# B&R Automation Studio project DemoCNC (part 2)

#### Variables.var - Local variables
```iecst
VAR
	deviceName : STRING[20] := 'CNC_PrgDir'; (*file device of the CNC programs (FileDevice of the axes group program feature, Config_4)*)
	shareParam : STRING[200] := '/SIP=192.0.2.20 /PROTOCOL=cifs /SHARE=GCode /USER=Controller /PASSWORD=change-me'; (*network share holding the CNC programs (HMI PC) - example values : set the address and the account of your PC*)
	step : USINT := 0;
	fbDevLink : DevLink;
	retryTimer : TON;
	linked : BOOL := FALSE; (*TRUE = the program folder is available*)
	linkStatus : UINT := 0; (*status of the last failed link, 0 = none*)
	sysError : UDINT := 0; (*FileIoGetSysError of the last failed link*)
END_VAR
```

### Package Logical/Motion - Manual axis moves, handwheel, path trace

### Program Logical/Motion/AxisManual (IEC) - Manual axis moves : jog, position move, single-axis commands

#### Init.st - Init code
```iecst
PROGRAM _INIT

	gEquipment.Output.Status.MoveComplete := TRUE;

	FOR i := 0 TO AX_LAST DO
		gAxis[i].Input.Parameter.JogSpeed := 50;
	END_FOR;

	(* static axis references : index 0 = X, 1 = Y, 2 = Z *)
	fbAxisInfo[AX_X].Axis := ADR(gAxis_X);
	fbAxisInfo[AX_Y].Axis := ADR(gAxis_Y);
	fbAxisInfo[AX_Z].Axis := ADR(gAxis_Z);

	fbAxisStatus[AX_X].Axis := ADR(gAxis_X);
	fbAxisStatus[AX_Y].Axis := ADR(gAxis_Y);
	fbAxisStatus[AX_Z].Axis := ADR(gAxis_Z);

	fbAxisPosition[AX_X].Axis := ADR(gAxis_X);
	fbAxisPosition[AX_Y].Axis := ADR(gAxis_Y);
	fbAxisPosition[AX_Z].Axis := ADR(gAxis_Z);

	fbAxisVelocity[AX_X].Axis := ADR(gAxis_X);
	fbAxisVelocity[AX_Y].Axis := ADR(gAxis_Y);
	fbAxisVelocity[AX_Z].Axis := ADR(gAxis_Z);

	fbAxisTorque[AX_X].Axis := ADR(gAxis_X);
	fbAxisTorque[AX_Y].Axis := ADR(gAxis_Y);
	fbAxisTorque[AX_Z].Axis := ADR(gAxis_Z);

	fbMoveAbs[AX_X].Axis := ADR(gAxis_X);
	fbMoveAbs[AX_Y].Axis := ADR(gAxis_Y);
	fbMoveAbs[AX_Z].Axis := ADR(gAxis_Z);

	fbMoveAdd[AX_X].Axis := ADR(gAxis_X);
	fbMoveAdd[AX_Y].Axis := ADR(gAxis_Y);
	fbMoveAdd[AX_Z].Axis := ADR(gAxis_Z);

	fbJog[AX_X].Axis := ADR(gAxis_X);
	fbJog[AX_Y].Axis := ADR(gAxis_Y);
	fbJog[AX_Z].Axis := ADR(gAxis_Z);

	fbStop[AX_X].Axis := ADR(gAxis_X);
	fbStop[AX_Y].Axis := ADR(gAxis_Y);
	fbStop[AX_Z].Axis := ADR(gAxis_Z);

	fbHalt[AX_X].Axis := ADR(gAxis_X);
	fbHalt[AX_Y].Axis := ADR(gAxis_Y);
	fbHalt[AX_Z].Axis := ADR(gAxis_Z);

	fbReset[AX_X].Axis := ADR(gAxis_X);
	fbReset[AX_Y].Axis := ADR(gAxis_Y);
	fbReset[AX_Z].Axis := ADR(gAxis_Z);

	fbAxisError[AX_X].Axis := ADR(gAxis_X);
	fbAxisError[AX_Y].Axis := ADR(gAxis_Y);
	fbAxisError[AX_Z].Axis := ADR(gAxis_Z);

	fbPower[AX_X].Axis := ADR(gAxis_X);
	fbPower[AX_Y].Axis := ADR(gAxis_Y);
	fbPower[AX_Z].Axis := ADR(gAxis_Z);

	fbHome[AX_X].Axis := ADR(gAxis_X);
	fbHome[AX_Y].Axis := ADR(gAxis_Y);
	fbHome[AX_Z].Axis := ADR(gAxis_Z);

	FOR i := 0 TO AX_LAST DO
		fbAxisInfo[i].Enable := TRUE;
		fbAxisStatus[i].Enable := TRUE;
		fbAxisPosition[i].Enable := TRUE;
		fbAxisVelocity[i].Enable := TRUE;
		fbAxisTorque[i].Enable := TRUE;
		fbAxisError[i].Enable := TRUE;

		fbJog[i].Acceleration := DEFAULT_ACC;
		fbJog[i].Deceleration := DEFAULT_DEC;
		fbMoveAbs[i].Acceleration := DEFAULT_ACC;
		fbMoveAbs[i].Deceleration := DEFAULT_DEC;
		fbMoveAdd[i].Acceleration := DEFAULT_ACC;
		fbMoveAdd[i].Deceleration := DEFAULT_DEC;
		fbStop[i].Deceleration := DEFAULT_DEC;
		fbHalt[i].Deceleration := DEFAULT_DEC;
	END_FOR

END_PROGRAM
```

#### Cyclic.st - Cyclic code
```iecst
PROGRAM _CYCLIC

	(* drive adapter PVs (Global.var) : referenced here so they are allocated on the target *)
	gDS402_X;
	gDS402_Y;
	gDS402_Z;

	(* copy the mappMotion position limits into gAxis[].Input.Parameter.SoftwareLimits* once after startup *)
	IF NOT cfgLimitLoaded THEN
		fbAxCfg.Name := cfgAxisName[cfgAxIdx];
		fbAxCfg.DataType := mcCFG_AX_MOVE_LIM;
		fbAxCfg.DataAddress := ADR(axMoveLim);
		fbAxCfg.Mode := mcPCM_LOAD;
		fbAxCfg.Execute := TRUE;
		fbAxCfg();

		IF fbAxCfg.Done OR fbAxCfg.Error THEN
			cfgLimitErrorID[cfgAxIdx] := fbAxCfg.ErrorID;
			IF fbAxCfg.Done THEN
				gAxis[cfgAxIdx].Input.Parameter.SoftwareLimitsNeg := LREAL_TO_DINT(axMoveLim.MovementLimits.Internal.Position.LowerLimit);
				gAxis[cfgAxIdx].Input.Parameter.SoftwareLimitsPos := LREAL_TO_DINT(axMoveLim.MovementLimits.Internal.Position.UpperLimit);
			END_IF
			fbAxCfg.Execute := FALSE;
			fbAxCfg();
			cfgAxIdx := cfgAxIdx + 1;
			cfgLimitLoaded := cfgAxIdx > AX_LAST;
		END_IF
	END_IF

	Torque_X := fbAxisTorque[AX_X].Torque;
	Torque_Y := fbAxisTorque[AX_Y].Torque;
	Torque_Z := fbAxisTorque[AX_Z].Torque;

	(* absolute positions are meaningless before homing *)
	allHomed := fbAxisInfo[AX_X].IsHomed AND fbAxisInfo[AX_Y].IsHomed AND fbAxisInfo[AX_Z].IsHomed;

	(* position move request of this scan : accepted or dropped below, reported by act_MoveResult *)
	moveReq := gEquipment.Input.Command.ManualMove;
	moveAccepted := FALSE;

	IF NOT DI_MPG_Jog_Enable AND gEquipment.Input.CncCommand = E_ACT_IDLE AND NOT gEquipment.Output.State.Move AND NOT DI_Auto AND NOT gEquipment.Output.Status.EmergencyStop THEN

		IF NOT allHomed THEN
			gEquipment.Input.Command.ManualMove := FALSE;
		END_IF

		IF gEquipment.Input.Command.ManualMove THEN
			gEquipment.Input.Command.ManualMove := FALSE;
			gEquipment.Output.Status.MoveComplete := FALSE;
			moveStep := 0;
			moveAccepted := TRUE;
		END_IF

		act_Jog;
	ELSE
		gEquipment.Output.Status.ManualMove := FALSE;
		gEquipment.Input.Command.ManualMove := FALSE; (* never run a stale move request later *)
	END_IF

	moveStepIn := moveStep;
	act_MovePosition;
	act_MoveResult; (* result to the HMI (gManualMoveResult) - reporting only *)

	(* per-axis POWER / HOME only while the CNC is idle *)
	cncIdle := gEquipment.Output.Status.CurrentAction = E_ACT_IDLE AND NOT gEquipment.Output.Status.ProgramActive;

	(* screen jog (Axis_JOG_POSITIVE / NEGATIVE) only in manual mode, without the handwheel and while no CNC command runs.
	   MOVE_ADDITIVE (one step) is not gated : the HMI uses it in auto mode too.
	   Not ProgramActive (cncIdle) : the axes group reports MoveActive for a cycle when a single axis starts to move, so every
	   jog would be dropped right after its start. A program only runs in auto mode, which NOT DI_Auto already keeps out *)
	jogAllowed := NOT DI_Auto AND NOT DI_MPG_Jog_Enable AND gEquipment.Output.Status.CurrentAction = E_ACT_IDLE;

	(* per-axis power is held by fbPower (Axis_POWER). E-stop and group servo off take the axes back *)
	IF gEquipment.Output.Status.EmergencyStop OR gEquipment.Output.Status.CurrentAction = E_ACT_POWER_OFF THEN
		FOR i := 0 TO AX_LAST BY 1 DO
			axisPowerReq[i] := FALSE;
		END_FOR
	END_IF

	(* jog watchdog : an HMI that changes gJogAlive while it jogs (every 0.1 s) gets the jog stopped when the value
	   stands still for 0.5 s (HMI hung, connection lost). An HMI that never changes it is not watched *)
	jogAny := jogPosActive[AX_X] OR jogNegActive[AX_X] OR jogPosActive[AX_Y] OR jogNegActive[AX_Y] OR jogPosActive[AX_Z] OR jogNegActive[AX_Z];
	IF NOT jogAny THEN
		jogAliveArmed := FALSE;
		jogAlivePrev := gJogAlive;
	ELSIF gJogAlive <> jogAlivePrev THEN
		jogAlivePrev := gJogAlive;
		jogAliveArmed := TRUE;
		jogAliveTimer(IN := FALSE); (* restart *)
	END_IF
	jogAliveTimer(IN := jogAny AND jogAliveArmed, PT := T#500ms);
	IF jogAliveTimer.Q THEN
		FOR i := 0 TO AX_LAST BY 1 DO
			jogPosActive[i] := FALSE;
			jogNegActive[i] := FALSE;
		END_FOR
		jogAliveArmed := FALSE;
	END_IF

	(* ---------- per-axis command handling ---------- *)
	FOR i := 0 TO AX_LAST BY 1 DO

		(* E-stop : stop whatever runs, accept only STOP / RESET *)
		IF gEquipment.Output.Status.EmergencyStop THEN
			IF gAxis[i].Input.Command.Command <> Axis_STOP AND gAxis[i].Input.Command.Command <> Axis_RESET THEN
				gAxis[i].Input.Command.Command := Axis_IDLE;
			END_IF
			IF (command[i] <> Axis_IDLE AND command[i] <> Axis_STOP AND command[i] <> Axis_RESET) OR jogPosActive[i] OR jogNegActive[i] THEN
				command[i] := Axis_STOP;
				commandStep[i] := 0;
			END_IF
		END_IF

		IF command[i] <> gAxis[i].Input.Command.Command AND command[i] = Axis_IDLE THEN
			gAxis[i].Output.State.Command := gAxis[i].Input.Command.Command;
			command[i] := gAxis[i].Input.Command.Command;
			gAxis[i].Input.Command.Command := Axis_IDLE;
			commandStep[i] := 0;
		ELSIF gAxis[i].Input.Command.Command = Axis_HALT AND command[i] <> Axis_IDLE THEN
			command[i] := gAxis[i].Input.Command.Command;
			gAxis[i].Input.Command.Command := Axis_IDLE;
			commandStep[i] := 0;
		ELSIF gAxis[i].Input.Command.Command = Axis_STOP AND command[i] <> Axis_IDLE THEN
			command[i] := gAxis[i].Input.Command.Command;
			gAxis[i].Input.Command.Command := Axis_IDLE;
			commandStep[i] := 0;
		END_IF

		(* a HALT / STOP ends a running position move (act_MovePosition never sends them itself) *)
		IF (command[i] = Axis_HALT OR command[i] = Axis_STOP) AND commandStep[i] = 0 AND moveStep < 100 THEN
			moveStep := 100;
		END_IF

		CASE command[i] OF
			Axis_IDLE:
				IF fbAxisInfo[i].IsHomed THEN
					gAxis[i].Output.State.Status := 1;
				ELSE
					gAxis[i].Output.State.Status := 0;
				END_IF

				gAxis[i].Output.State.Home := fbAxisInfo[i].IsHomed;

				(* keep jog active state while jogging (command returns to IDLE, motion continues) *)
				IF jogPosActive[i] OR jogNegActive[i] THEN
					gAxis[i].Output.State.Status := 2;
				END_IF

			Axis_HALT:
				CASE commandStep[i] OF
					0:
						IF (jogPosActive[i] OR jogNegActive[i]) AND NOT fbMoveAbs[i].Busy AND NOT fbMoveAdd[i].Busy AND NOT fbHome[i].Busy THEN
							(* jog only : the jog FB brakes by itself (Deceleration) when its request drops. MC_Halt would abort it,
							   and an aborted jog FB took no new jog until it was switched off and on *)
							jogPosActive[i] := FALSE;
							jogNegActive[i] := FALSE;
							fbMoveAbs[i].Execute := FALSE; (* not busy - released as in the MC_Halt path *)
							fbMoveAdd[i].Execute := FALSE;
							fbHome[i].Execute := FALSE;
							settleTimer[i](IN := FALSE);
							commandStep[i] := 2;
						ELSE
							jogPosActive[i] := FALSE;
							jogNegActive[i] := FALSE;
							fbMoveAbs[i].Execute := FALSE; (* release aborted moves so the next one gets a rising edge *)
							fbMoveAdd[i].Execute := FALSE;
							fbHome[i].Execute := FALSE;
							fbHalt[i].Execute := TRUE;
							settleTimer[i](IN := FALSE);
							commandStep[i] := 1;
						END_IF
					1:
						IF fbHalt[i].Done OR fbHalt[i].CommandAborted OR fbHalt[i].Error THEN
							fbHalt[i].Execute := FALSE;
							IF fbAxisStatus[i].StandStill OR fbAxisStatus[i].ErrorStop OR fbAxisStatus[i].Disabled THEN
								command[i] := Axis_IDLE;
							ELSE
								commandStep[i] := 2; (* status not yet standstill (read before the FB finished) *)
							END_IF
						END_IF
					2: (* wait for standstill (at most 2 s), then the channel is free again *)
						settleTimer[i](IN := TRUE, PT := T#2s);
						IF fbAxisStatus[i].StandStill OR fbAxisStatus[i].ErrorStop OR fbAxisStatus[i].Disabled OR settleTimer[i].Q THEN
							settleTimer[i](IN := FALSE);
							command[i] := Axis_IDLE;
						END_IF
				END_CASE

			Axis_HOME:
				(* single-axis homing with the homing settings of the axis configuration.
				   Group homing (Z first, then XY) is HOME / INIT in gEquipment.Input.CncCommand *)
				CASE commandStep[i] OF
					0:
						IF NOT cncIdle OR gEquipment.Output.Status.EmergencyStop OR NOT fbAxisInfo[i].PowerOn THEN
							command[i] := Axis_IDLE; (* rejected *)
						ELSE
							jogPosActive[i] := FALSE;
							jogNegActive[i] := FALSE;
							fbHome[i].HomingMode := mcHOMING_DEFAULT;
							fbHome[i].Execute := TRUE;
							gAxis[i].Output.State.Status := 2;
							commandStep[i] := 1;
						END_IF
					1:
						IF fbHome[i].Done OR fbHome[i].Error OR fbHome[i].CommandAborted THEN
							fbHome[i].Execute := FALSE;
							command[i] := Axis_IDLE;
						END_IF
				END_CASE

			Axis_POWER:
				(* gAxis[i].Input.Parameter.Power : TRUE = on, FALSE = off *)
				CASE commandStep[i] OF
					0:
						IF NOT cncIdle OR (gAxis[i].Input.Parameter.Power AND gEquipment.Output.Status.EmergencyStop) THEN
							command[i] := Axis_IDLE; (* rejected *)
						ELSIF gAxis[i].Input.Parameter.Power THEN
							axisPowerReq[i] := TRUE;
							commandStep[i] := 10;
						ELSIF NOT (fbAxisStatus[i].StandStill OR fbAxisStatus[i].Disabled OR fbAxisStatus[i].ErrorStop) THEN
							command[i] := Axis_IDLE; (* rejected : axis moving *)
						ELSE
							(* MC_Power switches off only on a falling Enable : take the axis first, then release it *)
							axisPowerReq[i] := TRUE;
							commandStep[i] := 20;
						END_IF
					10: (* on *)
						IF fbPower[i].Status OR fbPower[i].Error THEN
							command[i] := Axis_IDLE;
						END_IF
					20: (* off *)
						IF fbPower[i].Status OR fbPower[i].Error THEN
							axisPowerReq[i] := FALSE;
							commandStep[i] := 21;
						END_IF
					21:
						IF NOT fbAxisInfo[i].PowerOn OR fbPower[i].Error THEN
							command[i] := Axis_IDLE;
						END_IF
				END_CASE

			Axis_JOG_NEGATIVE:
				CASE commandStep[i] OF
					0:
						IF gAxis[i].Input.Parameter.JogSpeed = 0 THEN
							gAxis[i].Input.Parameter.JogSpeed := 50;
						END_IF

						IF NOT jogAllowed THEN
							command[i] := Axis_IDLE; (* rejected : auto mode, handwheel or CNC busy *)
						ELSIF jogFault[i] THEN
							jogFault[i] := FALSE; (* jog FB back on this scan - the jog request waits until it is ready (step 2) *)
							settleTimer[i](IN := FALSE);
							commandStep[i] := 2;
						ELSE
							gAxis[i].Output.State.JogNegative := TRUE;
							jogNegActive[i] := TRUE;
							jogPosActive[i] := FALSE;
							gAxis[i].Output.State.Status := 2;
							commandStep[i] := 1;
						END_IF
					1:
						command[i] := Axis_IDLE;
						commandStep[i] := 0;
					2: (* a request set before the FB reports Ready is not seen - the jog did not start *)
						settleTimer[i](IN := TRUE, PT := T#1s);
						IF fbJog[i].Ready OR settleTimer[i].Q THEN
							settleTimer[i](IN := FALSE);
							gAxis[i].Output.State.JogNegative := TRUE;
							jogNegActive[i] := TRUE;
							jogPosActive[i] := FALSE;
							gAxis[i].Output.State.Status := 2;
							commandStep[i] := 1;
						END_IF
				END_CASE

			Axis_JOG_POSITIVE:
				CASE commandStep[i] OF
					0:
						IF gAxis[i].Input.Parameter.JogSpeed = 0 THEN
							gAxis[i].Input.Parameter.JogSpeed := 50;
						END_IF

						IF NOT jogAllowed THEN
							command[i] := Axis_IDLE; (* rejected : auto mode, handwheel or CNC busy *)
						ELSIF jogFault[i] THEN
							jogFault[i] := FALSE; (* jog FB back on this scan - the jog request waits until it is ready (step 2) *)
							settleTimer[i](IN := FALSE);
							commandStep[i] := 2;
						ELSE
							gAxis[i].Output.State.JogPositive := TRUE;
							jogPosActive[i] := TRUE;
							jogNegActive[i] := FALSE;
							gAxis[i].Output.State.Status := 2;
							commandStep[i] := 1;
						END_IF
					1:
						command[i] := Axis_IDLE;
						commandStep[i] := 0;
					2: (* a request set before the FB reports Ready is not seen - the jog did not start *)
						settleTimer[i](IN := TRUE, PT := T#1s);
						IF fbJog[i].Ready OR settleTimer[i].Q THEN
							settleTimer[i](IN := FALSE);
							gAxis[i].Output.State.JogPositive := TRUE;
							jogPosActive[i] := TRUE;
							jogNegActive[i] := FALSE;
							gAxis[i].Output.State.Status := 2;
							commandStep[i] := 1;
						END_IF
				END_CASE

			Axis_MOVE_ABSOLUTE:
				CASE commandStep[i] OF
					0:
						IF NOT fbAxisInfo[i].IsHomed THEN
							(* absolute target without homing : reject *)
							command[i] := Axis_IDLE;
						ELSE
							fbMoveAbs[i].Position := gAxis[i].Input.Parameter.Position;
							fbMoveAbs[i].Velocity := gAxis[i].Input.Parameter.Speed; (* [mm/s] *)
							gAxis[i].Output.State.Status := 2;
							fbMoveAbs[i].Execute := TRUE;
							commandStep[i] := 1;
						END_IF
					1:
						IF fbMoveAbs[i].Done THEN
							fbMoveAbs[i].Execute := FALSE;
							command[i] := Axis_IDLE;
							commandStep[i] := 0;
						ELSIF fbMoveAbs[i].CommandAborted OR fbMoveAbs[i].Error THEN
							fbMoveAbs[i].Execute := FALSE;
							command[i] := Axis_IDLE;
							commandStep[i] := 0;
						END_IF
				END_CASE

			Axis_MOVE_ADDITIVE:
				CASE commandStep[i] OF
					0:
						gAxis[i].Output.State.Status := 2;
						fbMoveAdd[i].Distance := gAxis[i].Input.Parameter.Distance;
						fbMoveAdd[i].Velocity := gAxis[i].Input.Parameter.Speed;
						fbMoveAdd[i].Execute := TRUE;
						settleTimer[i](IN := FALSE);
						commandStep[i] := 1;
					1:
						IF fbMoveAdd[i].Done OR fbMoveAdd[i].CommandAborted OR fbMoveAdd[i].Error THEN
							fbMoveAdd[i].Execute := FALSE;
							IF fbAxisStatus[i].StandStill OR fbAxisStatus[i].ErrorStop OR fbAxisStatus[i].Disabled THEN
								command[i] := Axis_IDLE;
							ELSE
								commandStep[i] := 2; (* status not yet standstill (read before the FB finished) *)
							END_IF
						END_IF
					2: (* wait for standstill (at most 2 s), then the channel is free again *)
						settleTimer[i](IN := TRUE, PT := T#2s);
						IF fbAxisStatus[i].StandStill OR fbAxisStatus[i].ErrorStop OR fbAxisStatus[i].Disabled OR settleTimer[i].Q THEN
							settleTimer[i](IN := FALSE);
							command[i] := Axis_IDLE;
						END_IF
				END_CASE

			Axis_RESET:
				CASE commandStep[i] OF
					0:
						fbReset[i].Execute := TRUE;
						commandStep[i] := 1;
					1:
						IF fbReset[i].Done OR fbReset[i].Error THEN
							(* release even if the error remains - Output.State.Error shows it, a new RESET can be sent *)
							fbReset[i].Execute := FALSE;
							command[i] := Axis_IDLE;
						END_IF
				END_CASE

			Axis_STOP:
				CASE commandStep[i] OF
					0:
						jogPosActive[i] := FALSE;
						jogNegActive[i] := FALSE;
						fbMoveAbs[i].Execute := FALSE; (* release aborted moves so the next one gets a rising edge *)
						fbMoveAdd[i].Execute := FALSE;
						fbHome[i].Execute := FALSE;
						fbStop[i].Execute := TRUE;
						settleTimer[i](IN := FALSE);
						commandStep[i] := 1;
					1:
						IF fbStop[i].Done OR fbStop[i].Error THEN
							fbStop[i].Execute := FALSE;
							IF fbAxisStatus[i].StandStill OR fbAxisStatus[i].ErrorStop OR fbAxisStatus[i].Disabled THEN
								command[i] := Axis_IDLE;
							ELSE
								commandStep[i] := 2; (* MC_Stop holds the axis in Stopping until Execute falls *)
							END_IF
						END_IF
					2: (* wait for standstill (at most 2 s), then the channel is free again *)
						settleTimer[i](IN := TRUE, PT := T#2s);
						IF fbAxisStatus[i].StandStill OR fbAxisStatus[i].ErrorStop OR fbAxisStatus[i].Disabled OR settleTimer[i].Q THEN
							settleTimer[i](IN := FALSE);
							command[i] := Axis_IDLE;
						END_IF
				END_CASE

			ELSE
				(* Axis_MOVE_VELOCITY / unknown : not implemented - release so the axis channel is not locked *)
				command[i] := Axis_IDLE;
		END_CASE

		(* no jog during an E-stop *)
		IF gEquipment.Output.Status.EmergencyStop THEN
			jogPosActive[i] := FALSE;
			jogNegActive[i] := FALSE;
		END_IF

		(* auto mode, handwheel selected or a CNC command / program : a running screen jog stops too - the jog FB brakes
		   by itself (Deceleration) when its request drops, as on a HALT of a pure jog or the jog watchdog *)
		IF NOT jogAllowed THEN
			jogPosActive[i] := FALSE;
			jogNegActive[i] := FALSE;
		END_IF

		(* jog FB error or aborted (by MC_Halt / MC_Stop / a move / homing on the axis) : drop the jog and switch the FB off -
		   it leaves that state only on a falling Enable and took no new jog before (jog worked only now and then).
		   The next jog command switches it on again (no on/off toggling while the cause stays) *)
		IF fbJog[i].Error OR fbJog[i].CommandAborted THEN
			jogFault[i] := TRUE;
			jogPosActive[i] := FALSE;
			jogNegActive[i] := FALSE;
		END_IF

		(* while this axis jogs its speed follows the HMI (joystick tilt) - act_Jog copies it only while State.Move is FALSE *)
		IF (jogPosActive[i] OR jogNegActive[i]) AND gAxis[i].Input.Parameter.JogSpeed > 0 THEN
			JogSpeed[i] := gAxis[i].Input.Parameter.JogSpeed;
		END_IF

		(* jog FB : level controlled *)
		fbJog[i].Velocity := JogSpeed[i];
		fbJog[i].JogPositive := jogPosActive[i];
		fbJog[i].JogNegative := jogNegActive[i];
		fbJog[i].Enable := fbAxisInfo[i].PowerOn AND NOT jogFault[i];

		IF NOT jogPosActive[i] THEN
			gAxis[i].Output.State.JogPositive := FALSE;
		END_IF
		IF NOT jogNegActive[i] THEN
			gAxis[i].Output.State.JogNegative := FALSE;
		END_IF

		(* status to HMI - positions/velocities in measurement units [mm], [mm/s] *)
		gAxis[i].Output.State.Enable := fbAxisInfo[i].PowerOn;
		gAxis[i].Output.State.Position := fbAxisPosition[i].Position;
		gAxis[i].Output.State.Speed := fbAxisVelocity[i].Velocity;
		gAxis[i].Output.State.Error := fbAxisStatus[i].ErrorStop;
		gAxis[i].Output.State.ErrorID := DINT_TO_UDINT(fbAxisError[i].AxisErrorID);

		IF fbAxisStatus[i].ErrorStop THEN
			gAxis[i].Output.State.Status := 3;
		END_IF

		(* drive diagnosis to HMI (read only) - copies of the MC_ReadAxisInfo above, no new FB on the axis *)
		gDriveDiag[i].Valid := fbAxisInfo[i].Valid;
		gDriveDiag[i].CommReady := fbAxisInfo[i].CommunicationReady;
		gDriveDiag[i].ReadyForPowerOn := fbAxisInfo[i].ReadyForPowerOn;
		gDriveDiag[i].Warning := fbAxisInfo[i].AxisWarning;

		(* warning-level alarm (alarms.json exType 1) : filtered so one warning gives one alarm - display only, no reaction *)
		warnOnTimer[i](IN := gDriveDiag[i].Valid AND gDriveDiag[i].CommReady AND gDriveDiag[i].Warning, PT := T#500ms);
		warnHoldTimer[i](IN := warnOnTimer[i].Q, PT := T#2s);
		gDriveDiag[i].WarningAlarm := warnHoldTimer[i].Q;

		(* FB calls *)
		fbAxisInfo[i]();
		fbAxisStatus[i]();
		fbAxisPosition[i]();
		fbAxisVelocity[i]();
		fbAxisTorque[i]();
		fbAxisError[i]();
		fbMoveAbs[i]();
		fbMoveAdd[i]();
		fbJog[i]();
		fbStop[i]();
		fbHalt[i]();
		fbReset[i]();
		fbPower[i].Enable := axisPowerReq[i];
		fbPower[i]();
		fbHome[i]();

	END_FOR

END_PROGRAM
```

#### Exit.st - Exit code
```iecst
PROGRAM _EXIT
END_PROGRAM
```

#### Action_Jog.st - Jog action
```iecst
ACTION act_Jog:

	FOR i := 0 TO AX_LAST BY 1 DO
		JogSpeed[i] := gAxis[i].Input.Parameter.JogSpeed;
	END_FOR

END_ACTION
```

#### Action_MovePosition.st - Move position action
```iecst
ACTION act_MovePosition:

	(* abort on E-stop, axis error or lost homing - the wait steps below would never finish *)
	IF moveStep < 100 AND (NOT allHomed OR gEquipment.Output.Status.EmergencyStop OR gAxis[AX_X].Output.State.Error OR gAxis[AX_Y].Output.State.Error OR gAxis[AX_Z].Output.State.Error) THEN
		moveStep := 100;
	END_IF

	(* also end it when the machine leaves manual operation or an axis loses power, so it never
	   moves on by itself once the servo is back. A HALT / STOP of an axis ends it in Cyclic *)
	IF moveStep < 100 AND (DI_Auto OR DI_MPG_Jog_Enable OR gEquipment.Output.Status.CurrentAction <> E_ACT_IDLE OR
		NOT fbAxisInfo[AX_X].PowerOn OR NOT fbAxisInfo[AX_Y].PowerOn OR NOT fbAxisInfo[AX_Z].PowerOn) THEN
		moveStep := 100;
	END_IF

	CASE moveStep OF
		0:
			IF gAxis[AX_X].Input.Command.Command = Axis_IDLE AND gAxis[AX_Y].Input.Command.Command = Axis_IDLE AND gAxis[AX_Z].Input.Command.Command = Axis_IDLE THEN
				moveStep := 10;
			END_IF

		10: (* retract Z first *)
			gEquipment.Output.Status.ManualMove := TRUE;

			gAxis[AX_Z].Input.Parameter.Speed := gEquipment.Input.Parameter.SystemSpeed;
			gAxis[AX_Z].Input.Parameter.Position := 0;
			gAxis[AX_Z].Input.Command.Command := Axis_MOVE_ABSOLUTE;
			moveStep := 20;

		20:
			IF gAxis[AX_Z].Output.State.Status = 1 AND command[AX_Z] = Axis_IDLE AND fbAxisStatus[AX_Z].StandStill = TRUE THEN
				moveStep := 30;
			END_IF

		30: (* move X / Y *)
			gAxis[AX_X].Input.Parameter.Speed := gEquipment.Input.Parameter.SystemSpeed;
			gAxis[AX_X].Input.Parameter.Position := gEquipment.Input.Parameter.ManualPositon[0];
			gAxis[AX_X].Input.Command.Command := Axis_MOVE_ABSOLUTE;
			gAxis[AX_Y].Input.Parameter.Speed := gEquipment.Input.Parameter.SystemSpeed;
			gAxis[AX_Y].Input.Parameter.Position := gEquipment.Input.Parameter.ManualPositon[1];
			gAxis[AX_Y].Input.Command.Command := Axis_MOVE_ABSOLUTE;
			moveStep := 40;

		40:
			IF gAxis[AX_X].Output.State.Status = 1 AND gAxis[AX_Y].Output.State.Status = 1 AND
				command[AX_X] = Axis_IDLE AND command[AX_Y] = Axis_IDLE AND
				fbAxisStatus[AX_X].StandStill = TRUE AND fbAxisStatus[AX_Y].StandStill = TRUE AND fbAxisStatus[AX_Z].StandStill = TRUE THEN

				IF gEquipment.Input.Parameter.ManualSlowMove THEN
					gEquipment.Input.Parameter.ManualSlowMove := FALSE;
					moveStep := 45;
				ELSE
					moveStep := 50;
				END_IF
			END_IF

		45: (* approach : fast to (target - SlowMoveLength) *)
			gAxis[AX_Z].Input.Parameter.Speed := gEquipment.Input.Parameter.SystemSpeed;
			gAxis[AX_Z].Input.Parameter.Position := gEquipment.Input.Parameter.ManualPositon[2] - SlowMoveLength;
			gAxis[AX_Z].Input.Command.Command := Axis_MOVE_ABSOLUTE;
			moveStep := 46;

		46:
			IF gAxis[AX_Z].Output.State.Status = 1 AND command[AX_Z] = Axis_IDLE AND fbAxisStatus[AX_Z].StandStill = TRUE THEN
				moveStep := 47;
			END_IF

		47: (* slow final approach *)
			gAxis[AX_Z].Input.Parameter.Speed := gEquipment.Input.Parameter.SystemSpeed * SlowMoveVelocity / 100;
			gAxis[AX_Z].Input.Parameter.Position := gEquipment.Input.Parameter.ManualPositon[2];
			gAxis[AX_Z].Input.Command.Command := Axis_MOVE_ABSOLUTE;
			moveStep := 60;

		50:
			gAxis[AX_Z].Input.Parameter.Speed := gEquipment.Input.Parameter.SystemSpeed;
			gAxis[AX_Z].Input.Parameter.Position := gEquipment.Input.Parameter.ManualPositon[2];
			gAxis[AX_Z].Input.Command.Command := Axis_MOVE_ABSOLUTE;
			moveStep := 60;

		60:
			IF gAxis[AX_Z].Output.State.Status = 1 AND command[AX_Z] = Axis_IDLE AND fbAxisStatus[AX_Z].StandStill = TRUE THEN
				moveStep := 100;
			END_IF

		100:
			gEquipment.Output.Status.ManualMove := FALSE;
			gEquipment.Output.Status.MoveComplete := TRUE;
	END_CASE
END_ACTION
```

#### Action_MoveResult.st - Move position result action
```iecst
ACTION act_MoveResult:

	(* result of the position move (Input.Command.ManualMove) for the HMI : gManualMoveResult - reporting only, the move
	   (Cyclic acceptance, act_MovePosition) is not changed. Called right after act_MovePosition, so the checks below see the values it saw.
	   A refused request and a cancelled move are reported as such, not as arrived *)

	(* why act_MovePosition ends a running move in this scan - its two checks, MOVE_RSN_NONE = it does not *)
	IF gEquipment.Output.Status.EmergencyStop THEN
		moveEndReason := MOVE_RSN_ESTOP;
	ELSIF DI_Auto THEN
		moveEndReason := MOVE_RSN_AUTO;
	ELSIF DI_MPG_Jog_Enable THEN
		moveEndReason := MOVE_RSN_HANDWHEEL;
	ELSIF gEquipment.Output.Status.CurrentAction <> E_ACT_IDLE THEN
		moveEndReason := MOVE_RSN_CNC_BUSY;
	ELSIF gAxis[AX_X].Output.State.Error OR gAxis[AX_Y].Output.State.Error OR gAxis[AX_Z].Output.State.Error THEN
		moveEndReason := MOVE_RSN_AXIS_ERROR;
	ELSIF NOT fbAxisInfo[AX_X].PowerOn OR NOT fbAxisInfo[AX_Y].PowerOn OR NOT fbAxisInfo[AX_Z].PowerOn THEN
		moveEndReason := MOVE_RSN_SERVO_OFF;
	ELSIF NOT allHomed THEN
		moveEndReason := MOVE_RSN_NOT_HOMED;
	ELSE
		moveEndReason := MOVE_RSN_NONE;
	END_IF

	IF moveReq THEN
		(* a request was taken in this scan : Result / Reason now belong to request number Count *)
		gManualMoveResult.Count := gManualMoveResult.Count + 1;
		gManualMoveResult.Reason := MOVE_RSN_NONE;
		moveFailed := FALSE;

		IF NOT moveAccepted THEN
			(* dropped by the acceptance in Cyclic - its conditions in this order *)
			gManualMoveResult.Result := MOVE_RES_REFUSED;
			IF gEquipment.Output.Status.EmergencyStop THEN
				gManualMoveResult.Reason := MOVE_RSN_ESTOP;
			ELSIF DI_Auto THEN
				gManualMoveResult.Reason := MOVE_RSN_AUTO;
			ELSIF DI_MPG_Jog_Enable THEN
				gManualMoveResult.Reason := MOVE_RSN_HANDWHEEL;
			ELSIF gEquipment.Input.CncCommand <> E_ACT_IDLE THEN
				gManualMoveResult.Reason := MOVE_RSN_CNC_BUSY;
			ELSIF gEquipment.Output.State.Move THEN
				gManualMoveResult.Reason := MOVE_RSN_MOVING;
			ELSE
				gManualMoveResult.Reason := MOVE_RSN_NOT_HOMED; (* the only other case Cyclic drops it *)
			END_IF
		ELSIF moveStep >= 100 THEN
			(* accepted, but act_MovePosition ended it in the same scan (servo off, axis error, CNC command) : nothing moved *)
			gManualMoveResult.Result := MOVE_RES_REFUSED;
			gManualMoveResult.Reason := moveEndReason;
		ELSE
			gManualMoveResult.Result := MOVE_RES_RUNNING;
		END_IF

	ELSIF gManualMoveResult.Result = MOVE_RES_RUNNING THEN
		(* an absolute move of the sequence ended aborted or with an error : the sequence goes on, the target may not be reached.
		   The FB outputs are still set here - the axis step 1 in Cyclic releases them later in this scan *)
		FOR i := 0 TO AX_LAST BY 1 DO
			IF fbMoveAbs[i].CommandAborted OR fbMoveAbs[i].Error THEN
				moveFailed := TRUE;
			END_IF
		END_FOR

		IF moveStepIn >= 100 THEN
			(* ended between two scans : only the axis HALT / STOP check in Cyclic does that *)
			gManualMoveResult.Result := MOVE_RES_CANCELLED;
			gManualMoveResult.Reason := MOVE_RSN_AXIS_HALT;
		ELSIF moveStep >= 100 THEN
			IF moveEndReason <> MOVE_RSN_NONE THEN
				gManualMoveResult.Result := MOVE_RES_CANCELLED;
				gManualMoveResult.Reason := moveEndReason;
			ELSIF moveFailed THEN
				gManualMoveResult.Result := MOVE_RES_CANCELLED;
				gManualMoveResult.Reason := MOVE_RSN_STEP_FAILED;
			ELSE
				gManualMoveResult.Result := MOVE_RES_ARRIVED; (* step 60 : every step of the sequence done *)
			END_IF
		END_IF
	END_IF

END_ACTION
```

#### Variables.var - Local variables
```iecst
VAR CONSTANT
	DEFAULT_ACC : REAL := 500.0; (* [mm/s^2] - keep consistent with axis config MovementLimits *)
	DEFAULT_DEC : REAL := 500.0; (* [mm/s^2] *)
END_VAR
VAR
	i : INT := 0;
	command : ARRAY[0..2] OF AXIS_COMMAND;
	commandStep : ARRAY[0..2] OF SINT;
	moveStep : USINT := 100;
	JogSpeed : ARRAY[0..2] OF REAL;
	jogPosActive : ARRAY[0..2] OF BOOL := [3(FALSE)];
	jogNegActive : ARRAY[0..2] OF BOOL := [3(FALSE)];
	allHomed : BOOL := FALSE;
	cncIdle : BOOL := FALSE;
	axisPowerReq : ARRAY[0..2] OF BOOL := [3(FALSE)]; (*per-axis power held by fbPower (Axis_POWER)*)
	settleTimer : ARRAY[0..2] OF TON; (*HALT / STOP / MOVE_ADDITIVE step 2 : release the channel at the latest after this if the axis does not report standstill*)
	jogFault : ARRAY[0..2] OF BOOL := [3(FALSE)]; (*jog FB had an error : held off until the next jog command*)
	jogAllowed : BOOL := FALSE; (*screen jog (Axis_JOG_POSITIVE / NEGATIVE) taken and kept : manual mode, no handwheel, no CNC command (CurrentAction IDLE)*)
END_VAR
(*jog watchdog (gJogAlive from the HMI)*)
VAR
	jogAny : BOOL := FALSE; (*some axis is jogging*)
	jogAliveArmed : BOOL := FALSE; (*gJogAlive changed during this jog : the HMI is watched*)
	jogAlivePrev : UINT := 0;
	jogAliveTimer : TON; (*gJogAlive standing still while jogging*)
END_VAR
(*drive warning alarm filter (gDriveDiag[].WarningAlarm)*)
VAR
	warnOnTimer : ARRAY[0..2] OF TON; (*the drive warning must stand this long before WarningAlarm rises*)
	warnHoldTimer : ARRAY[0..2] OF TOF; (*WarningAlarm stays this long after the warning clears*)
END_VAR
(*position move result to the HMI (gManualMoveResult, act_MoveResult) - reporting only*)
VAR CONSTANT
	MOVE_RES_RUNNING : USINT := 1;
	MOVE_RES_ARRIVED : USINT := 2;
	MOVE_RES_REFUSED : USINT := 3;
	MOVE_RES_CANCELLED : USINT := 4; (*ended before the target, the reason says why*)
	MOVE_RSN_NONE : USINT := 0;
	MOVE_RSN_ESTOP : USINT := 1;
	MOVE_RSN_AUTO : USINT := 2;
	MOVE_RSN_HANDWHEEL : USINT := 3;
	MOVE_RSN_CNC_BUSY : USINT := 4;
	MOVE_RSN_MOVING : USINT := 5;
	MOVE_RSN_NOT_HOMED : USINT := 6;
	MOVE_RSN_SERVO_OFF : USINT := 7;
	MOVE_RSN_AXIS_ERROR : USINT := 8;
	MOVE_RSN_AXIS_HALT : USINT := 9;
	MOVE_RSN_STEP_FAILED : USINT := 10;
END_VAR
VAR
	moveReq : BOOL := FALSE; (*a ManualMove request was there at the start of this scan (Cyclic takes it in every case)*)
	moveAccepted : BOOL := FALSE; (*that request started the sequence*)
	moveStepIn : USINT := 100; (*moveStep before act_MovePosition of this scan*)
	moveEndReason : USINT := 0; (*why act_MovePosition ends a running move in this scan (its two checks), MOVE_RSN_NONE = it does not*)
	moveFailed : BOOL := FALSE; (*an absolute axis move of the running sequence ended aborted or with an error*)
END_VAR
(* mapp Motion axis FBs *)
VAR
	fbAxisInfo : ARRAY[0..2] OF MC_ReadAxisInfo;
	fbAxisStatus : ARRAY[0..2] OF MC_ReadStatus;
	fbAxisPosition : ARRAY[0..2] OF MC_ReadActualPosition;
	fbAxisVelocity : ARRAY[0..2] OF MC_ReadActualVelocity;
	fbAxisTorque : ARRAY[0..2] OF MC_ReadActualTorque;
	fbMoveAbs : ARRAY[0..2] OF MC_MoveAbsolute;
	fbMoveAdd : ARRAY[0..2] OF MC_MoveAdditive;
	fbJog : ARRAY[0..2] OF MC_BR_JogVelocity;
	fbStop : ARRAY[0..2] OF MC_Stop;
	fbHalt : ARRAY[0..2] OF MC_Halt;
	fbReset : ARRAY[0..2] OF MC_Reset;
	fbAxisError : ARRAY[0..2] OF MC_ReadAxisError;
	fbPower : ARRAY[0..2] OF MC_Power;
	fbHome : ARRAY[0..2] OF MC_Home;
END_VAR
(* software limits read once from the mappMotion axis config at startup, copied into gAxis[].Input.Parameter.SoftwareLimitsNeg / Pos *)
VAR
	fbAxCfg : MC_BR_ProcessConfig;
	axMoveLim : McCfgAxMoveLimType;
	cfgAxisName : ARRAY[0..2] OF STRING[32] := ['gAxis_X','gAxis_Y','gAxis_Z'];
	cfgAxIdx : USINT := 0;
	cfgLimitLoaded : BOOL := FALSE;
	cfgLimitErrorID : ARRAY[0..2] OF DINT; (*ErrorID of reading the limits of that axis, 0 = read. On an error the limits of that axis stay 0 : ZRef refuses, the handwheel stops at 0*)
END_VAR
```

### Program Logical/Motion/Handwheel (IEC) - Handwheel (MPG)

#### Init.st - Init code
```iecst
PROGRAM _INIT

	axisRef[AX_X] := ADR(gAxis_X);
	axisRef[AX_Y] := ADR(gAxis_Y);
	axisRef[AX_Z] := ADR(gAxis_Z);

	FOR i := 0 TO AX_LAST DO
		fbMpgMove[i].Axis := axisRef[i];
		fbMpgStop[i].Axis := axisRef[i];
		fbMpgPosition[i].Axis := axisRef[i];
		fbMpgStatus[i].Axis := axisRef[i];
		fbMpgPosition[i].Enable := TRUE;
		fbMpgStatus[i].Enable := TRUE;
		fbMpgMove[i].Acceleration := MPG_ACC;
		fbMpgMove[i].Deceleration := MPG_ACC;
		fbMpgStop[i].Deceleration := MPG_ACC;
	END_FOR

END_PROGRAM
```

#### Cyclic.st - Cyclic code
```iecst
PROGRAM _CYCLIC

	(* handwheel mode starts : every axis takes its reference again *)
	enableRise(CLK := DI_MPG_Jog_Enable);

	IF enableRise.Q THEN
		FOR i := 0 TO AX_LAST DO
			axisActive[i] := FALSE;
		END_FOR
	END_IF

	(* E-stop : stop the handwheel axis, drop the reference so the next use resyncs to the actual position *)
	emgTrig(CLK := gEquipment.Output.Status.EmergencyStop);

	IF emgTrig.Q THEN
		FOR i := 0 TO AX_LAST DO
			axisActive[i] := FALSE;
			movePending[i] := FALSE;
			fbMpgMove[i].Execute := FALSE;
			fbMpgStop[i].Execute := TRUE;
		END_FOR
	END_IF

	IF gEquipment.Input.CncCommand = E_ACT_IDLE AND NOT gEquipment.Output.State.Move AND NOT gEquipment.Output.Status.EmergencyStop THEN

		IF DI_MPG_AxisX THEN
			selectAxis := 1;
		ELSIF DI_MPG_AxisY THEN
			selectAxis := 2;
		ELSIF DI_MPG_AxisZ THEN
			selectAxis := 3;
		END_IF

		IF selectAxis > 0 THEN
			act_SelectAxis;
			act_SelectStep;

			IF counterReset THEN
				(* counter is being reset : resync so the jump to 0 is not counted as movement *)
				prevCounter := counterValue;
				counterSynced := FALSE;
			ELSE
				act_CountPulses;
			END_IF
		END_IF

		(* counter reset : one cycle pulse *)
		IF selectAxis > 0 AND counterReset THEN
			counterReset := FALSE;
		END_IF

		axisChange(CLK := selectAxis <> lastSelectAxis);

		IF axisChange.Q THEN
			lastSelectAxis := selectAxis;
			counterReset := TRUE;

			(* axis changed without passing through OFF : drop the previous axis reference *)
			FOR i := 0 TO AX_LAST DO
				axisActive[i] := FALSE;
				movePending[i] := FALSE;
				fbMpgMove[i].Execute := FALSE;
			END_FOR
			prevCounter := 0;
			counterSynced := FALSE;
		END_IF

		(* axis selector back to OFF : stop, reset the counter *)
		axisReleased(CLK := DI_MPG_AxisX OR DI_MPG_AxisY OR DI_MPG_AxisZ);

		IF axisReleased.Q THEN
			selectAxis := 0;
			counterReset := TRUE;
			prevCounter := 0;
			counterSynced := FALSE;
			FOR i := 0 TO AX_LAST DO
				axisActive[i] := FALSE;
				fbMpgStop[i].Execute := TRUE;
				movePending[i] := FALSE;
				fbMpgMove[i].Execute := FALSE;
			END_FOR
		END_IF

	END_IF

	(* release stop execute after done *)
	FOR i := 0 TO AX_LAST DO
		IF fbMpgStop[i].Execute AND (fbMpgStop[i].Done OR fbMpgStop[i].Error) THEN
			fbMpgStop[i].Execute := FALSE;
		END_IF
	END_FOR

	(* MC_MoveAbsolute retrigger : drop Execute one scan, re-arm with new target *)
	FOR i := 0 TO AX_LAST DO
		IF movePending[i] AND NOT fbMpgMove[i].Execute THEN
			fbMpgMove[i].Execute := TRUE;
			movePending[i] := FALSE;
		END_IF

		IF fbMpgMove[i].Execute AND (fbMpgMove[i].Done OR fbMpgMove[i].Error OR fbMpgMove[i].CommandAborted) THEN
			fbMpgMove[i].Execute := FALSE;
		END_IF

		fbMpgMove[i]();
		fbMpgStop[i]();
		fbMpgPosition[i]();
		fbMpgStatus[i]();
	END_FOR

END_PROGRAM
```

#### Exit.st - Exit code
```iecst
PROGRAM _EXIT
END_PROGRAM
```

#### Action_Handwheel.st - Handwheel actions
```iecst
(* selected axis (selectAxis 1..3 = X..Z) : stop the other axes, take the actual position as the start of the target once *)
ACTION act_SelectAxis:

	ax := selectAxis - 1;

	FOR i := 0 TO AX_LAST DO
		IF i <> ax AND NOT fbMpgStatus[i].StandStill THEN
			fbMpgStop[i].Execute := TRUE;
			axisActive[i] := FALSE;
		END_IF
	END_FOR

	IF NOT axisActive[ax] THEN
		axisActive[ax] := TRUE;
		target := fbMpgPosition[ax].Position;
	END_IF

	fbMpgMove[ax].Velocity := gAxis[ax].Input.Parameter.JogSpeed; (* [mm/s] *)

END_ACTION

(* step per detent from the x1 / x10 / x100 selector *)
ACTION act_SelectStep:

	IF DI_MPG_X1 THEN
		stepPerDetent := STEP_X1;
	ELSIF DI_MPG_X10 THEN
		stepPerDetent := STEP_X10;
	ELSIF DI_MPG_X100 THEN
		stepPerDetent := STEP_X100;
	END_IF

END_ACTION

(* counter change -> new target of the active axis, kept inside the software limits.
   The first change after a reset only synchronises the counter *)
ACTION act_CountPulses:

	delta := counterValue - prevCounter;

	IF delta <> 0 THEN

		IF NOT counterSynced THEN
			counterSynced := TRUE;
			prevCounter := counterValue;
			RETURN;
		END_IF

		FOR i := 0 TO AX_LAST DO
			IF axisActive[i] THEN
				target := target + DINT_TO_LREAL(delta) * stepPerDetent / COUNTS_PER_DETENT;
				IF delta > 0 THEN
					target := MIN(target, DINT_TO_LREAL(gAxis[i].Input.Parameter.SoftwareLimitsPos));
				ELSE
					target := MAX(target, DINT_TO_LREAL(gAxis[i].Input.Parameter.SoftwareLimitsNeg));
				END_IF
				fbMpgMove[i].Position := target;
				fbMpgMove[i].Execute := FALSE; (* drop -> re-armed next scan *)
				movePending[i] := TRUE;
			END_IF
		END_FOR

	END_IF

	prevCounter := counterValue;

END_ACTION
```

#### Variables.var - Local variables
```iecst
VAR CONSTANT
	STEP_X1 : LREAL := 0.01; (*[mm/detent] selector x1*)
	STEP_X10 : LREAL := 0.1; (*[mm/detent] selector x10*)
	STEP_X100 : LREAL := 1.0; (*[mm/detent] selector x100*)
	COUNTS_PER_DETENT : LREAL := 4.0; (*encoder counts per detent (quadrature x4)*)
	MPG_ACC : REAL := 500.0; (*[mm/s^2]*)
END_VAR
VAR
	selectAxis : USINT := 0; (*axis selected on the handwheel, 1..3 = X..Z, 0 = none*)
	lastSelectAxis : USINT := 0;
	ax : USINT; (*selectAxis - 1*)
	axisRef : ARRAY[0..2] OF UDINT; (*ADR of gAxis_X/Y/Z*)
	i : USINT;
	axisActive : ARRAY[0..2] OF BOOL; (*the axis follows the handwheel, target taken from its position*)
	target : LREAL; (*target position of the active axis [mm]*)
	stepPerDetent : LREAL;
	counterReset : BOOL; (*IoMap : %QX X20DC1176 Encoder01Reset*)
	counterValue : DINT; (*IoMap : %ID X20DC1176 Encoder01*)
	prevCounter : DINT;
	delta : DINT;
	counterSynced : BOOL; (*FALSE after a reset : the next counter change only synchronises*)
	movePending : ARRAY[0..2] OF BOOL;
	enableRise : R_TRIG;
	axisChange : R_TRIG;
	axisReleased : F_TRIG;
	emgTrig : R_TRIG;
END_VAR
(*mapp Motion FBs*)
VAR
	fbMpgMove : ARRAY[0..2] OF MC_MoveAbsolute;
	fbMpgStop : ARRAY[0..2] OF MC_Stop;
	fbMpgPosition : ARRAY[0..2] OF MC_ReadActualPosition;
	fbMpgStatus : ARRAY[0..2] OF MC_ReadStatus;
END_VAR
```

### Program Logical/Motion/RingBuffer (IEC) - Ring buffer of the axis path for the HMI 3D trace

#### Cyclic.st - Cyclic code
```iecst
(* Records axis positions, head on (discharge or laser), moving state, the laser power and the value of the
   active head into a ring buffer. Runs in Cyclic#1 (2ms), same task class as the motion programs. *)
PROGRAM _CYCLIC
	BufferX[Head] := gAxis[AX_X].Output.State.Position;
	BufferY[Head] := gAxis[AX_Y].Output.State.Position;
	BufferZ[Head] := gAxis[AX_Z].Output.State.Position;
	BufferHeadOn[Head] := gDispenser.Input.Command.Discharge OR gLaser.Input.Command.Emission;
	BufferMoving[Head] := gEquipment.Output.State.Move;
	BufferLaserPower[Head] := REAL_TO_USINT(LIMIT(0.0, gLaser.Output.State.Power, 100.0));
	(* value of the active head : the laser power for the laser - also while the head is not known (gActiveHead 0),
	   the laser is the only head with a value - and 0 for a head without a value (dispenser) *)
	IF gActiveHead = 0 OR gActiveHead = HEAD_LASER THEN
		BufferHeadValue[Head] := BufferLaserPower[Head];
	ELSE
		BufferHeadValue[Head] := 0;
	END_IF

	Head := Head + 1;
	IF Head >= RB_SIZE THEN
		Head := 0;
	END_IF
END_PROGRAM
```

#### Init.st - Init code
```iecst
PROGRAM _INIT
	Head := 0;
END_PROGRAM
```

#### Exit.st - Exit code
```iecst
PROGRAM _EXIT
END_PROGRAM
```

#### Variables.var - Local variables
```iecst
VAR CONSTANT
	RB_SIZE : UDINT := 500; (*number of samples: 500 * 2ms = 1s history.
	                          HMI polls every ~100ms - the buffer only bridges poll gaps.
	                          Kept small so the HMI reads stay fast and regular.*)
	RB_MAX : UDINT := 499; (*RB_SIZE - 1*)
END_VAR

VAR
	BufferX : ARRAY[0..RB_MAX] OF LREAL; (*X axis actual position [mm]*)
	BufferY : ARRAY[0..RB_MAX] OF LREAL; (*Y axis actual position [mm]*)
	BufferZ : ARRAY[0..RB_MAX] OF LREAL; (*Z axis actual position [mm]*)
	BufferHeadOn : ARRAY[0..RB_MAX] OF BOOL; (*TRUE while discharge or laser emission command is active*)
	BufferMoving : ARRAY[0..RB_MAX] OF BOOL; (*TRUE while the equipment is moving.
	                                           Sampled here so the HMI reads it on the same
	                                           time base as the positions - the subscription
	                                           value alone runs ahead of the buffered samples.*)
	BufferLaserPower : ARRAY[0..RB_MAX] OF USINT; (*laser power output [%] (gLaser.Output.State.Power, after corner compensation, 0 while off).
	                                                The HMI shades the 3D laser trace with it. One scan old - Laser runs after RingBuffer.*)
	BufferHeadValue : ARRAY[0..RB_MAX] OF USINT; (*value of the active head 0..100 (gActiveHead) for the HMI head plugins - laser : = BufferLaserPower
	                                               (also while gActiveHead is 0), dispenser : 0 (no value)*)
	Head : UDINT := 0; (*next write position, wraps at RB_SIZE*)
END_VAR
```

### Package Logical/Heads - Dispenser and laser head outputs

### Program Logical/Heads/Dispenser (IEC) - Dispenser discharge output

#### Cyclic.st - Cyclic code
```iecst
PROGRAM _CYCLIC

	(* mode change (auto <-> manual) : discharge off, both commands dropped *)
	toAuto(CLK := gEquipment.Output.Status.Mode);
	toManual(CLK := gEquipment.Output.Status.Mode);
	IF toAuto.Q OR toManual.Q THEN
		gDispenser.Input.Command.Discharge := FALSE;
		gDispenser.Input.Command.Manual := FALSE;
		DO_Dispenser_Start := FALSE;
	END_IF

	(* auto : M41 / M42 (Command.Discharge, driven by Main), manual : Command.Manual from the HMI *)
	IF gEquipment.Output.Status.Mode THEN
		command := gDispenser.Input.Command.Discharge;
	ELSE
		command := gDispenser.Input.Command.Manual;
	END_IF

	(* on with the rising edge (not in dry run), off with the falling edge *)
	commandOn(CLK := command);
	commandOff(CLK := command);

	IF commandOn.Q AND NOT gEquipment.Input.Parameter.DryRun THEN
		DO_Dispenser_Start := TRUE;
	ELSIF commandOff.Q THEN
		DO_Dispenser_Start := FALSE;
	END_IF

	gDispenser.Output.State.Discharge := DO_Dispenser_Start;

END_PROGRAM
```

#### Init.st - Init code
```iecst
PROGRAM _INIT

END_PROGRAM
```

#### Exit.st - Exit code
```iecst
PROGRAM _EXIT
	DO_Dispenser_Start := FALSE;
END_PROGRAM
```

#### Variables.var - Local variables
```iecst
VAR
	toAuto : R_TRIG;
	toManual : F_TRIG;
	command : BOOL; (*discharge command of the current mode*)
	commandOn : R_TRIG;
	commandOff : F_TRIG;
END_VAR
```

### Program Logical/Heads/Laser (IEC) - PWM laser output

#### Cyclic.st - Cyclic code
```iecst
PROGRAM _CYCLIC

	autoOn(CLK := gEquipment.Output.Status.Mode);
	autoOff(CLK := gEquipment.Output.Status.Mode);

	IF autoOn.Q OR autoOff.Q THEN
		gLaser.Input.Command.Manual := FALSE;
	END_IF

	(* laser allowed : not in dry run or E-stop *)
	supplyOn := NOT (gEquipment.Input.Parameter.DryRun OR gEquipment.Output.Status.EmergencyStop);

	(* emission : level controlled - auto : M61 / M62 (Emission is driven by Main), manual : Command.Manual *)
	IF gEquipment.Output.Status.Mode THEN
		emissionOn := gLaser.Input.Command.Emission;
	ELSE
		emissionOn := gLaser.Input.Command.Manual;
	END_IF
	emissionOn := emissionOn AND supplyOn;

	(* X20DO8331 DO02 (on/off laser output) is held off : the PWM laser on X20DO4332-1 is switched on and off by its duty below *)
	DO_Laser_Power := FALSE;

	(* power [%] : manual test power, else LaserPower of the program, else the auto power *)
	IF NOT gEquipment.Output.Status.Mode THEN
		power := gLaser.Input.Parameter.ManualPower;
	ELSIF C_LaserPower >= 0.0 THEN
		power := C_LaserPower;
	ELSE
		power := gLaser.Input.Parameter.Power;
	END_IF

	(* corner compensation : power x actual / programmed path velocity, so a slower path (corners, feed override) does not burn deeper *)
	fbPathInfo.Enable := gLaser.Input.Parameter.SpeedScale AND gEquipment.Output.Status.ProgramActive;
	fbPathInfo();
	speedRatio := 1.0;
	IF fbPathInfo.Valid AND gEquipment.Output.Status.Mode AND fbPathInfo.PathInfo.ProgrammedPathVelocity > 0.0 THEN
		speedRatio := LIMIT(LIMIT(0.0, gLaser.Input.Parameter.MinSpeedRatio, 100.0) / 100.0,
			fbPathInfo.PathInfo.CurrentPathVelocity / fbPathInfo.PathInfo.ProgrammedPathVelocity, 1.0);
	END_IF
	power := LIMIT(0.0, power * speedRatio, 100.0);

	(* PWM : power 0..100 % -> duty DutyMin..DutyMax, duty 0 while off or at power 0 *)
	IF emissionOn AND power > 0.0 THEN
		duty := LIMIT(0.0, gLaser.Input.Parameter.DutyMin + (gLaser.Input.Parameter.DutyMax - gLaser.Input.Parameter.DutyMin) * power / 100.0, 100.0);
	ELSE
		duty := 0.0;
		power := 0.0;
	END_IF

	PWM_Laser_Duty := REAL_TO_INT(duty * 327.67);
	PWM_Laser_Period := MAX(gLaser.Input.Parameter.PwmPeriod, 1000); (* 0 would switch PWM off in the module, below 1000 us is not allowed *)
	DO_Laser_On := emissionOn AND PWM_Laser_Duty > 0;

	gLaser.Output.State.Emission := DO_Laser_On;
	gLaser.Output.State.Power := power;
	gLaser.Output.State.Duty := duty;

END_PROGRAM
```

#### Init.st - Init code
```iecst
PROGRAM _INIT

	(* gLaser is not RETAIN : the HMI writes the head table values when they differ from these.
	   Until then the laser stays dark (power 0) - a program can still set LaserPower. *)
	gLaser.Input.Parameter.Power := 0.0;
	gLaser.Input.Parameter.ManualPower := 0.0;
	gLaser.Input.Parameter.DutyMin := 0.0;
	gLaser.Input.Parameter.DutyMax := 100.0;
	gLaser.Input.Parameter.PwmPeriod := 1000; (* 1 kHz *)
	gLaser.Input.Parameter.SpeedScale := FALSE;
	gLaser.Input.Parameter.MinSpeedRatio := 20.0;

	fbPathInfo.AxesGroup := ADR(gCncXYZ);

	DO_Laser_Power := FALSE;
	DO_Laser_On := FALSE;
	PWM_Laser_Duty := 0;

END_PROGRAM
```

#### Exit.st - Exit code
```iecst
PROGRAM _EXIT

	DO_Laser_Power := FALSE;
	DO_Laser_On := FALSE;
	PWM_Laser_Duty := 0;

	fbPathInfo.Enable := FALSE;
	fbPathInfo();

END_PROGRAM
```

#### Variables.var - Local variables
```iecst
VAR
	autoOn : R_TRIG;
	autoOff : F_TRIG;
	fbPathInfo : MC_BR_PathInfo; (*actual / programmed path velocity for the corner compensation*)
	supplyOn : BOOL := FALSE; (*laser allowed (no dry run, heavy alarm, E-stop)*)
	emissionOn : BOOL := FALSE; (*laser commanded on (auto Emission / manual) and supply on*)
	power : REAL := 0.0; (*power [%] after the source selection and the corner compensation*)
	speedRatio : REAL := 1.0; (*actual / programmed path velocity, limited to MinSpeedRatio..1*)
	duty : REAL := 0.0; (*PWM duty [%]*)
END_VAR
```
